DATA_BLOCK "GDB_RecoveryStamp"
{ S7_Optimized_Access := 'TRUE' }
VERSION : 0.1
NON_RETAIN
VAR
    Data {ExternalAccessible := 'False'; ExternalVisible := 'False'; ExternalWritable := 'False'} : DTL;
END_VAR
BEGIN
END_DATA_BLOCK
